{region 'Documentation'}
(*!
<summary>Render a quoted diagnostic preview with at most AssertionValueLength output bytes.
Printable ASCII is retained; other code units become byte 16#D7 without expansion.</summary>
<description>
Zero terminates the input. Quotes and backslashes remain literal. Shortening reserves
space for enclosing quotes and an ellipsis; the default limit retains 35 code units.
Rendering is lossy and does not alter the compared input or its result.
</description>
*)
{endregion}
FUNCTION INTERNAL CreateAssertionTextValue_String : STRING(GVL_Constants.AssertionValueLength) //! Bounded diagnostic aid; not a lossless representation for subsequent comparison.
VAR_INPUT
    Value : STRING(GVL_Constants.MessageLength); //! Text to preview; zero terminates the input.
END_VAR
VAR
    Text : STRING(GVL_Constants.AssertionValueLength);
    CharacterIndex : INT;
    CopyLength : INT;
    Code : BYTE;
    Shortened : BOOL;
END_VAR
VAR CONSTANT
    Quote : STRING(1) := '$'';
    Ellipsis : STRING(3) := '...';
    QuoteLength : INT := 2;
    EllipsisLength : INT := 3;
    FirstPrintableAscii : BYTE := 16#20;
    LastPrintableAscii : BYTE := 16#7E;
    ReplacementByte : BYTE := 16#D7;
END_VAR

CopyLength := UINT_TO_INT(GVL_Constants.AssertionValueLength) - QuoteLength;
// SA0175: Bounded diagnostic code-unit rendering; each unsupported unit becomes one byte.
{analysis -175}
Shortened := TRUE;
FOR CharacterIndex := 0 TO CopyLength DO
    IF Value[CharacterIndex] = 0 THEN
        CopyLength := CharacterIndex;
        Shortened := FALSE;
        EXIT;
    END_IF;
END_FOR;
IF Shortened THEN
    CopyLength := CopyLength - EllipsisLength;
END_IF;

FOR CharacterIndex := 0 TO CopyLength - 1 DO
    Code := Value[CharacterIndex];
    IF (Code >= FirstPrintableAscii) AND (Code <= LastPrintableAscii) THEN
        Text[CharacterIndex] := Code;
    ELSE
        Text[CharacterIndex] := ReplacementByte;
    END_IF;
END_FOR;
Text[CopyLength] := 0;
{analysis +175}

IF Shortened THEN
    Text := CONCAT(Text, Ellipsis);
END_IF;
CreateAssertionTextValue_String := CONCAT(Quote, Text);
CreateAssertionTextValue_String := CONCAT(CreateAssertionTextValue_String, Quote);

END_FUNCTION

(* stored: Version 1.1.0.1
   POU CreateAssertionTextValue_String: Id {f3ee0d93-3f4e-4348-9924-baa2fdd4a505}, SpecialFunc None *)
